(*
SPDX-FileCopyrightText: © 2026 Oleksandr Tiutyk <trofimich@gmail.com>
SPDX-License-Identifier: MIT
License: https://opensource.org/license/mit
*)

(*!
<summary>Provides fluent assertions on a copied LREAL value.</summary>
<description>
Copies actual into persistent instance storage before the entry method returns; literals and expression
results therefore remain valid throughout the immediate chain. Owns no heap allocation or pointed-to resource.
The message prefixes every failure until the next preparation. Finish one chain before starting another on
the owning Assertions provider. Use only from the owning test callback on one task, without reentry.
Obtain this context from the owning provider; direct unprepared use is unsupported.
Expected arguments use the declared IEC type; ordinary compiler conversions happen before comparison.
This context does not depend on another assertion context.
Object metadata is available before preparation; inherited equality compares instance identity.
Equality and inclusive ordering accept a finite nonnegative LREAL tolerance, default zero. Strict ordering
has no tolerance. Core canonical NaN, infinity and signed-zero rules apply; unequal nonfinite values are
never close. Invalid tolerance records failure without throwing. Tolerance belongs only to that method call.
Inclusive ordering also accepts equality from Core ordering under the target's floating configuration;
exact ToBe and NotToBe still compare canonical bits when tolerance is zero.
</description>
*)

{attribute 'no_explicit_call' := 'do not call this function block directly'}
FUNCTION_BLOCK LongRealAssertionContext EXTENDS TOF_Core.Object
VAR_STAT
	{attribute 'hide'}
	_ClassName : STRING := __POUNAME();
END_VAR
VAR
	_Actual : LREAL;
	_TestCase : ITestCase;
	_Message : WSTRING(255);
END_VAR

(*!
<summary>Provides the implementation class name.</summary>
<description>
Borrowed read-only reference to compiler-initialized storage, valid throughout the instance lifetime.
Do not modify the returned reference; no ownership is transferred.
</description>
*)
{attribute 'monitoring' := 'call'}
PROPERTY ClassName : REFERENCE TO STRING
GET
ClassName REF= _ClassName;
END_GET
END_PROPERTY

(*!
<summary>Asserts that the actual value is strictly greater than expected.</summary>
<description>
Records failure without interrupting the callback; preserves the message for the rest of the chain.
</description>
<param name="expected">Expected value converted by the compiler to LREAL.</param>
*)
METHOD FINAL IsGreaterThan : REFERENCE TO LongRealAssertionContext
VAR_INPUT
	expected : LREAL;
END_VAR
VAR
	actualBits : ULINT;
	expectedBits : ULINT;
	comparison : TOF_Core.COMPARISON_RESULT;
END_VAR
actualBits := TestServices.GetCanonicalLongRealBits(value := _Actual);
expectedBits := TestServices.GetCanonicalLongRealBits(value := expected);

comparison := TestServices.CompareFloatingValues(
	actualBits := actualBits,
	expectedBits := expectedBits
);

IF comparison <> TOF_Core.COMPARISON_RESULT.FIRST_GREATER_THAN_SECOND THEN
	failComparison(
		expected := expected,
		expectation := "Expected value > "
	);
END_IF

IsGreaterThan REF= THIS^;
END_METHOD

(*!
<summary>Asserts that the actual value meets the inclusive lower boundary.</summary>
<description>
Records failure without interrupting the callback; preserves the message for the rest of the chain.
Uses the canonical floating policy shared by the typed contexts, matching Core semantics, and absolute tolerance.
Invalid tolerance records failure before comparison. The default zero does not affect later assertions in this chain.
</description>
<param name="expected">Expected value converted by the compiler to LREAL.</param>
<param name="tolerance">Finite nonnegative absolute distance for this call only; default zero.</param>
*)
METHOD FINAL IsGreaterThanOrEquals : REFERENCE TO LongRealAssertionContext
VAR_INPUT
	expected : LREAL;
	tolerance : LREAL := LREAL#0.0;
END_VAR
VAR
	actualBits : ULINT;
	expectedBits : ULINT;
	comparison : TOF_Core.COMPARISON_RESULT;
	isSatisfied : BOOL;
END_VAR
IF NOT TestServices.IsValidFloatingTolerance(tolerance := tolerance) THEN
	TestServices.ReportAssertionFailure(
		testCase := _TestCase,
		message := _Message,
		sourceClassName := ClassName,
		defaultMessage := "Expected a finite nonnegative comparison tolerance"
	);
	IsGreaterThanOrEquals REF= THIS^;
	RETURN;
END_IF

actualBits := TestServices.GetCanonicalLongRealBits(value := _Actual);
expectedBits := TestServices.GetCanonicalLongRealBits(value := expected);

comparison := TestServices.CompareFloatingValues(
	actualBits := actualBits,
	expectedBits := expectedBits
);

isSatisfied := (comparison = TOF_Core.COMPARISON_RESULT.FIRST_GREATER_THAN_SECOND)
	OR_ELSE (comparison = TOF_Core.COMPARISON_RESULT.FIRST_EQUAL_TO_SECOND)
	OR_ELSE TestServices.AreFloatingValuesWithinTolerance(
		actualBits := actualBits,
		expectedBits := expectedBits,
		tolerance := tolerance
	);

IF NOT isSatisfied THEN
	failComparison(
		expected := expected,
		expectation := "Expected value >= ",
		toleranceText := TOF_Core.WideStrings.Concat255(", tolerance: ", TO_WSTRING(tolerance))
	);
END_IF

IsGreaterThanOrEquals REF= THIS^;
END_METHOD

(*!
<summary>Asserts that the actual value is strictly less than expected.</summary>
<description>
Records failure without interrupting the callback; preserves the message for the rest of the chain.
</description>
<param name="expected">Expected value converted by the compiler to LREAL.</param>
*)
METHOD FINAL IsLessThan : REFERENCE TO LongRealAssertionContext
VAR_INPUT
	expected : LREAL;
END_VAR
VAR
	actualBits : ULINT;
	expectedBits : ULINT;
	comparison : TOF_Core.COMPARISON_RESULT;
END_VAR
actualBits := TestServices.GetCanonicalLongRealBits(value := _Actual);
expectedBits := TestServices.GetCanonicalLongRealBits(value := expected);

comparison := TestServices.CompareFloatingValues(
	actualBits := actualBits,
	expectedBits := expectedBits
);

IF comparison <> TOF_Core.COMPARISON_RESULT.FIRST_LESS_THAN_SECOND THEN
	failComparison(
		expected := expected,
		expectation := "Expected value < "
	);
END_IF

IsLessThan REF= THIS^;
END_METHOD

(*!
<summary>Asserts that the actual value meets the inclusive upper boundary.</summary>
<description>
Records failure without interrupting the callback; preserves the message for the rest of the chain.
Uses the canonical floating policy shared by the typed contexts, matching Core semantics, and absolute tolerance.
Invalid tolerance records failure before comparison. The default zero does not affect later assertions in this chain.
</description>
<param name="expected">Expected value converted by the compiler to LREAL.</param>
<param name="tolerance">Finite nonnegative absolute distance for this call only; default zero.</param>
*)
METHOD FINAL IsLessThanOrEquals : REFERENCE TO LongRealAssertionContext
VAR_INPUT
	expected : LREAL;
	tolerance : LREAL := LREAL#0.0;
END_VAR
VAR
	actualBits : ULINT;
	expectedBits : ULINT;
	comparison : TOF_Core.COMPARISON_RESULT;
	isSatisfied : BOOL;
END_VAR
IF NOT TestServices.IsValidFloatingTolerance(tolerance := tolerance) THEN
	TestServices.ReportAssertionFailure(
		testCase := _TestCase,
		message := _Message,
		sourceClassName := ClassName,
		defaultMessage := "Expected a finite nonnegative comparison tolerance"
	);
	IsLessThanOrEquals REF= THIS^;
	RETURN;
END_IF

actualBits := TestServices.GetCanonicalLongRealBits(value := _Actual);
expectedBits := TestServices.GetCanonicalLongRealBits(value := expected);

comparison := TestServices.CompareFloatingValues(
	actualBits := actualBits,
	expectedBits := expectedBits
);

isSatisfied := (comparison = TOF_Core.COMPARISON_RESULT.FIRST_LESS_THAN_SECOND)
	OR_ELSE (comparison = TOF_Core.COMPARISON_RESULT.FIRST_EQUAL_TO_SECOND)
	OR_ELSE TestServices.AreFloatingValuesWithinTolerance(
		actualBits := actualBits,
		expectedBits := expectedBits,
		tolerance := tolerance
	);

IF NOT isSatisfied THEN
	failComparison(
		expected := expected,
		expectation := "Expected value <= ",
		toleranceText := TOF_Core.WideStrings.Concat255(", tolerance: ", TO_WSTRING(tolerance))
	);
END_IF

IsLessThanOrEquals REF= THIS^;
END_METHOD

(*!
<summary>Provides the library namespace.</summary>
<description>
Borrowed read-only reference to the compiler-initialized namespace, valid throughout the instance lifetime.
Do not modify the returned reference; no ownership is transferred.
</description>
*)
{attribute 'monitoring' := 'call'}
PROPERTY NamespaceName : REFERENCE TO STRING
GET
NamespaceName REF= CurrentNamespace.Name;
END_GET
END_PROPERTY

(*!
<summary>Asserts inequality with the expected value.</summary>
<description>
Records failure without interrupting the callback; preserves the message for the rest of the chain.
Uses the canonical floating policy shared by the typed contexts, matching Core semantics, and absolute tolerance.
Invalid tolerance records failure before comparison. The default zero does not affect later assertions in this chain.
</description>
<param name="expected">Expected value converted by the compiler to LREAL.</param>
<param name="tolerance">Finite nonnegative absolute distance for this call only; default zero.</param>
*)
METHOD FINAL NotToBe : REFERENCE TO LongRealAssertionContext
VAR_INPUT
	expected : LREAL;
	tolerance : LREAL := LREAL#0.0;
END_VAR
VAR
	actualBits : ULINT;
	expectedBits : ULINT;
	areEqual : BOOL;
END_VAR
IF NOT TestServices.IsValidFloatingTolerance(tolerance := tolerance) THEN
	TestServices.ReportAssertionFailure(
		testCase := _TestCase,
		message := _Message,
		sourceClassName := ClassName,
		defaultMessage := "Expected a finite nonnegative comparison tolerance"
	);
	NotToBe REF= THIS^;
	RETURN;
END_IF

actualBits := TestServices.GetCanonicalLongRealBits(value := _Actual);
expectedBits := TestServices.GetCanonicalLongRealBits(value := expected);

areEqual := TestServices.AreFloatingValuesWithinTolerance(
	actualBits := actualBits,
	expectedBits := expectedBits,
	tolerance := tolerance
);

IF areEqual THEN
	failComparison(
		expected := expected,
		expectation := "Expected value not to be: ",
		toleranceText := TOF_Core.WideStrings.Concat255(", tolerance: ", TO_WSTRING(tolerance))
	);
END_IF

NotToBe REF= THIS^;
END_METHOD

(*!
<summary>Copies the actual operand and replaces the chain-wide message.</summary>
<description>
Called by the owning Assertions provider after it verifies the running test case.
No pointer to this method's input storage is retained. The receiver is borrowed until the next preparation;
the owning provider keeps it alive throughout the immediate chain.
</description>
<param name="actual">Value copied into this context.</param>
<param name="testCase">Borrowed failure receiver for the immediate chain.</param>
<param name="message">Copied diagnostic prefix, including empty to clear the previous prefix.</param>
*)
METHOD INTERNAL FINAL Prepare
VAR_INPUT
	actual : LREAL;
	testCase : ITestCase;
	message : WSTRING(255);
END_VAR
_Actual := actual;
_TestCase := testCase;
_Message := message;
END_METHOD

(*!
<summary>Reports the byte size of this concrete instance.</summary>
<description>
Includes inline fields and nested instances, but excludes separately allocated payloads.
Obtaining the size does not transfer ownership or validate an arbitrary address.
</description>
*)
{attribute 'monitoring' := 'call'}
PROPERTY SelfSize : ULINT
GET
SelfSize := XSIZEOF(THIS^);
END_GET
END_PROPERTY

(*!
<summary>Asserts equality with the expected value.</summary>
<description>
Records failure without interrupting the callback; preserves the message for the rest of the chain.
Uses the canonical floating policy shared by the typed contexts, matching Core semantics, and absolute tolerance.
Invalid tolerance records failure before comparison. The default zero does not affect later assertions in this chain.
</description>
<param name="expected">Expected value converted by the compiler to LREAL.</param>
<param name="tolerance">Finite nonnegative absolute distance for this call only; default zero.</param>
*)
METHOD FINAL ToBe : REFERENCE TO LongRealAssertionContext
VAR_INPUT
	expected : LREAL;
	tolerance : LREAL := LREAL#0.0;
END_VAR
VAR
	actualBits : ULINT;
	expectedBits : ULINT;
	areEqual : BOOL;
END_VAR
IF NOT TestServices.IsValidFloatingTolerance(tolerance := tolerance) THEN
	TestServices.ReportAssertionFailure(
		testCase := _TestCase,
		message := _Message,
		sourceClassName := ClassName,
		defaultMessage := "Expected a finite nonnegative comparison tolerance"
	);
	ToBe REF= THIS^;
	RETURN;
END_IF

actualBits := TestServices.GetCanonicalLongRealBits(value := _Actual);
expectedBits := TestServices.GetCanonicalLongRealBits(value := expected);

areEqual := TestServices.AreFloatingValuesWithinTolerance(
	actualBits := actualBits,
	expectedBits := expectedBits,
	tolerance := tolerance
);

IF NOT areEqual THEN
	failComparison(
		expected := expected,
		expectation := "Expected: ",
		toleranceText := TOF_Core.WideStrings.Concat255(", tolerance: ", TO_WSTRING(tolerance))
	);
END_IF

ToBe REF= THIS^;
END_METHOD

(*!
<summary>Formats a failed typed predicate and reports it with the chain message.</summary>
<description>
Does not change operands or chain state. The receiver retains its first failure. Reporting exceptions
propagate to the enclosing test callback handler; an unprepared receiver is a configuration error.
</description>
<param name="expected">Typed expected operand used only for this diagnostic.</param>
<param name="expectation">Prefix identifying the failed predicate.</param>
<param name="toleranceText">Optional call-local tolerance suffix; empty for strict ordering.</param>
*)
METHOD PRIVATE failComparison
VAR_INPUT
	expected : LREAL;
	expectation : WSTRING(40);
	toleranceText : WSTRING(80) := "";
END_VAR
VAR
	actualText : WSTRING(255);
	expectedText : WSTRING(255);
	diagnostic : TOF_Core.ERROR_MESSAGE;
END_VAR
actualText := TO_WSTRING(_Actual);
expectedText := TO_WSTRING(expected);

diagnostic := TOF_Core.WideStrings.Concat255(
	expectation,
	expectedText,
	", but was: ",
	actualText,
	toleranceText
);

TestServices.ReportAssertionFailure(
	testCase := _TestCase,
	message := _Message,
	sourceClassName := ClassName,
	defaultMessage := diagnostic
);
END_METHOD

END_FUNCTION_BLOCK

(* stored: Version 1.1.0.1
   POU LongRealAssertionContext: Id {a5f54457-4793-4012-a7f2-fe2d2bb49a23}, SpecialFunc None
   Folder Service methods: Id {60bb22b7-9019-4407-a992-b8d991af433f}
   Property ClassName: Id {d92388fc-43c0-4125-951b-e64ffb9529e6}
   Get Get: Id {834cff07-bc82-4c2e-9a1b-8f9c75d3ac01}
   Method IsGreaterThan: Id {46064e09-845a-415a-bbb7-940fa7dde37a}
   Method IsGreaterThanOrEquals: Id {ec90c7ea-22ea-4213-8767-23ca8fcc6653}
   Method IsLessThan: Id {cec3440d-e2f1-46ce-b803-9f377f740ffe}
   Method IsLessThanOrEquals: Id {a9274064-b06c-43eb-9317-1279610fc832}
   Property NamespaceName: Id {ed66e186-7060-4f64-a203-6b0019d2bdef}
   Get Get: Id {3bde8c19-48a1-425c-98e9-98d05095c1a4}
   Method NotToBe: Id {8716d711-b266-429b-b1bf-e5a00ca7dcd5}
   Method Prepare: Id {8f48c619-8751-4e6a-a790-5110e63d0486}
   Property SelfSize: Id {61e093c0-ef22-4098-b215-a451879deccd}
   Get Get: Id {45d19d2b-bf06-413b-9b96-7a7c8318412e}
   Method ToBe: Id {3ca43e1e-71fa-470e-93da-043250423ec9}
   Method failComparison: Id {5331a9e3-4dab-4f38-8502-81a51f9f945c} *)
